(* IEC 61131-3 sources: plc-vscode/tests/st/all/rusty/tests/integration/data/empty_proj/src, 1 file *)

(* ---- mainProg.st ---- *)
PROGRAM mainProg
VAR
x : DINT;
END_VAR

x := 1;
END_PROGRAM
